FUNCTION_BLOCK AD_TO_AD2 (* Composite FB for convert unidirectional AD to bidirectional AD2 *)
  (* Standard: 61499-2; Function: AD_IN publishes its value onto the outgoing (EO1) side of AD2_BIDIR. Whatever AD2_BIDIR receives on its incoming (EI1) side is forwarded out again as a plain unidirectional signal via AD_OUT.; Description: Copyright (c) 2026 HR Agrartechnik GmbH This program and the accompanying materials are made available under the terms of the Eclipse Public License 2.0 which is available at https://www.eclipse.org/legal/epl-2.0/ SPDX-License-Identifier: EPL-2.0 *)
  (* Version 1.0, 2026-10-13, Franz Höpfinger, HR Agrartechnik GmbH, Initial Version - Konvertierungsfamilie vervollstaendigt (analog zu AUI_TO_AUI2/AR_TO_AR2/AB_TO_AB2). *)
  PACKAGE adapter::conversion::bidirectional;
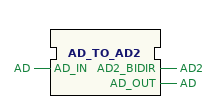
  SOCKETS
    AD_IN : adapter::types::unidirectional::AD; (* Adapter Input: unidirectional source *)
  END_SOCKETS
  PLUGS
    AD2_BIDIR : adapter::types::bidirectional::AD2; (* Adapter Output: bidirectional tap, outgoing side driven by AD_IN, incoming side forwarded to AD_OUT *)
    AD_OUT : adapter::types::unidirectional::AD; (* Adapter Output: mirrors AD2_BIDIR's incoming (request) side *)
  END_PLUGS
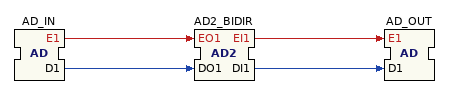
  EVENT_CONNECTIONS
    AD_IN.E1 TO AD2_BIDIR.EO1;
    AD2_BIDIR.EI1 TO AD_OUT.E1;
  END_CONNECTIONS
  DATA_CONNECTIONS
    AD_IN.D1 TO AD2_BIDIR.DO1;
    AD2_BIDIR.DI1 TO AD_OUT.D1;
  END_CONNECTIONS
END_FUNCTION_BLOCK
